// TIA Portal V20 export
VAR_GLOBAL   // PLC tag table "PLC-A3-AI"
   RESERVE_AI AT %IW64 : Int;
END_VAR
